(* IEC 61131-3 sources: Jacob-Formschaumtechnik-ISEL-CNC-Retrofit/twincat/PLC/src/6_Interfaces, 5 files *)

(* ---- Alarm_Catalog.st ---- *)
(* Meldekatalog: Slot-Nummer = Index in aCond von FB_AlarmList.
   Klassen siehe E_FaultClass. Texte und Abhilfe stehen in docs/Meldeliste.md (HMI-Thread). *)
TYPE E_AlarmSlot :
(
    SafetyOpen := 0,
    DoorOpen := 1,
    AirPressureLow := 2,
    ExtractionFault := 3,
    SpindleFuFault := 4,
    SpindlePtcTrip := 5,
    SpindleNoFeedback := 6,
    SpindleLockedSetup := 7,
    AxisDriveFault := 8,
    AxisFollowingErr := 9,
    HwLimitHit := 10,
    FieldbusLost := 11,
    HomingLost := 12,
    HmiLinkLost := 13,
    ParamMismatch := 14
) INT;
END_TYPE

(* ---- ST_HmiCmd.st ---- *)
(* HMI -> SPS. Die HMI fordert nur an. Alle Verriegelungen liegen in der SPS. *)
TYPE ST_HmiCmd :
STRUCT
    nHeartbeat      : UINT;    (* Lebenszeichen, wird von der HMI hochgezaehlt *)
    eModeRequest    : E_OpMode;
    bStart          : BOOL;    (* Impuls *)
    bHold           : BOOL;    (* Impuls, Vorschubhalt *)
    bAbort          : BOOL;    (* Impuls *)
    bAck            : BOOL;    (* Impuls, Meldungen quittieren, Wiederanlauf *)
    bJogPlus        : BOOL;    (* gehalten, nur mit Heartbeat *)
    bJogMinus       : BOOL;
    nJogAxis        : USINT;   (* 1=X, 2=Y, 3=Z *)
    bJogRapid       : BOOL;
    bSpindleOn      : BOOL;    (* nur Hand *)
    bSpindleCcw     : BOOL;
    rSpindleSetRpm  : REAL;    (* 1/min *)
    bExtraction     : BOOL;
    bBlowAir        : BOOL;
    bVacuum         : BOOL;
    bHomeRequest    : BOOL;    (* Impuls *)
    bToolChangeDone : BOOL;    (* Impuls, Quittung manueller Werkzeugwechsel *)
END_STRUCT
END_TYPE

(* ---- ST_HmiSts.st ---- *)
(* SPS -> HMI. CNC-Werte (Achspositionen, Overrides, Werkzeug-/Nullpunkttabelle) liest die HMI
   direkt aus der CNC (TF5310 Datenmodell), nicht ueber diese Struktur. *)
TYPE ST_HmiSts :
STRUCT
    eMode           : E_OpMode;
    eState          : E_MachState;
    bSafetyOk       : BOOL;
    bDrivesEnabled  : BOOL;
    bAllHomed       : BOOL;
    bHmiLinkOk      : BOOL;    (* Heartbeat der HMI wird ueberwacht *)
    bSpindleRunning : BOOL;
    rSpindleActRpm  : REAL;
    bExtractionOn   : BOOL;
    bBlowAirOn      : BOOL;
    bVacuumOn       : BOOL;
    bToolChangeReq  : BOOL;    (* Aufforderung am Panel *)
    nToolChangeNo   : UINT;
    nTopAlarmId     : INT;     (* hoechste aktive Meldung, 0 = keine *)
    eTopAlarmClass  : E_FaultClass;
    nActiveAlarms   : UINT;
    nMachineId      : UINT;    (* aus Maschinenparametern, z. B. 1 fuer M1 *)
    sSwVersion      : STRING(15);
    dwOperatingSec  : UDINT;   (* Betriebssekunden, fuer Wartungsanzeige *)
    dwSpindleSec    : UDINT;
END_STRUCT
END_TYPE

(* ---- ST_MachineParams.st ---- *)
(* Maschinenparameter. Je Maschine eine Datei in config/, geladen beim Start.
   Werte in config/M1.json mit [Annahme] gekennzeichnet, solange nicht bestaetigt. *)
TYPE ST_MachineParams :
STRUCT
    nMachineId        : UINT;
    sSwVersionExpected: STRING(15);
    nNumAxes          : USINT;             (* NC-Achsen ohne Spindel *)
    rSpindleMaxRpm    : REAL;              (* 16600 fuer VKH63/26-90T *)
    rSpindleMinRpm    : REAL;
    rSpindleVoltMax   : REAL;              (* 10.0 V entspricht rSpindleMaxRpm *)
    tSpindleRunUp     : TIME;              (* Wartezeit nach Start bis Drehzahl erreicht *)
    tSpindleStandstill: TIME;              (* Auslaufzeit bis Stillstand gemeldet *)
    tHmiTimeout       : TIME;              (* Heartbeat-Ausfall -> Tippen stoppt *)
    tFeedbackTimeout  : TIME;              (* Rueckmeldung Ventil/Spindel *)
    bAirMonitoring    : BOOL;
    bHasToolChanger   : BOOL;
END_STRUCT
END_TYPE

(* ---- Types_Common.st ---- *)
(* P-016 Gemeinsame Typen. Alle Maschinen M1 bis M4 nutzen diesen Stand. *)

TYPE E_OpMode :
(
    Hand  := 0,   (* Tippen, Handrad, Referenzieren *)
    Auto  := 1,   (* Programmbetrieb *)
    Setup := 2    (* Einrichten/Test: Spindel gesperrt, Einzelsatz moeglich *)
) INT;
END_TYPE

TYPE E_MachState :
(
    Stopped     := 0,  (* Antriebe aus, kein Fehler *)
    Idle        := 1,  (* Antriebe bereit, kein Programm *)
    Execute     := 2,  (* Programm laeuft *)
    Held        := 3,  (* Vorschubhalt, Programm fortsetzbar *)
    Aborted     := 4,  (* Programm abgebrochen, Reset noetig *)
    EStop       := 5,  (* Sicherheitskreis offen *)
    Fault       := 6   (* Fehler R3/R4 aktiv, Quittierung noetig *)
) INT;
END_TYPE

(* Fehlerreaktionsklassen, siehe docs/Architektur_Sicherheit.md *)
TYPE E_FaultClass :
(
    R0_Info     := 0,  (* nur anzeigen *)
    R1_Warning  := 1,  (* anzeigen, Betrieb laeuft weiter *)
    R2_FeedHold := 2,  (* gefuehrter Vorschubhalt, fortsetzbar *)
    R3_Abort    := 3,  (* gefuehrter Halt, Spindel aus, Programm beendet *)
    R4_DrivesOff := 4  (* Reglerfreigabe weg, Referenz verloren *)
) INT;
END_TYPE

TYPE E_AlarmId :
(
    None              := 0,
    SafetyOpen        := 100,  (* Sicherheitskreis offen / NOT-HALT *)
    DoorOpen          := 101,
    AirPressureLow    := 110,
    ExtractionFault   := 120,
    SpindleFuFault    := 200,
    SpindlePtcTrip    := 201,
    SpindleNoFeedback := 202,
    SpindleLockedSetup:= 203,
    AxisDriveFault    := 300,
    AxisFollowingErr  := 301,
    HwLimitHit        := 302,
    FieldbusLost      := 310,
    HomingLost        := 320,
    ParamMismatch     := 900   (* Maschinen-ID oder Version passt nicht *)
) INT;
END_TYPE

(* Eine Meldung aus der Meldeliste *)
TYPE ST_Alarm :
STRUCT
    eId    : E_AlarmId;
    eClass : E_FaultClass;
    bActive : BOOL;
    bAcked  : BOOL;
END_STRUCT
END_TYPE
